FUNCTION_BLOCK FB_AdmittanceController
VAR_INPUT
	
END_VAR
VAR_OUTPUT
END_VAR
VAR
END_VAR

END_FUNCTION_BLOCK

(* stored: Version 1.1.0.1, ProductVersion 3.1.4024.15
   POU FB_AdmittanceController: Id {697ed3a3-8819-4187-8c2f-568655b4914b}, SpecialFunc None *)
